(* IEC 61131-3 sources: plc-vscode/tests/st/test-ready/rusty/tests/lit/single/polymorphism/properties, 4 files *)

(* ---- alternating_accessor_overrides.st ---- *)
// RUN: (%COMPILE %s && %RUN) | %CHECK %s
// Scenario: Three-level POU chain C → B → A. B overrides only the getter (adds 1000),
// C overrides only the setter (adds 2000). Dispatch through POINTER TO A should resolve
// each accessor independently to the most-derived override:
//   A → (A.get, A.set)
//   B → (B.get, A.set)
//   C → (B.get, C.set)

FUNCTION_BLOCK A
    VAR
        _val : DINT := 10;
    END_VAR

    PROPERTY_GET value: DINT
        value := _val;
    END_PROPERTY

    PROPERTY_SET value: DINT
        _val := value;
    END_PROPERTY

    METHOD printValue
        printf('value=%d$N', value);
    END_METHOD

    METHOD setValue
        VAR_INPUT x : DINT; END_VAR
        value := x;
    END_METHOD
END_FUNCTION_BLOCK

FUNCTION_BLOCK B EXTENDS A
    // Override only getter — adds 1000
    PROPERTY_GET value: DINT
        value := _val + 1000;
    END_PROPERTY
END_FUNCTION_BLOCK

FUNCTION_BLOCK C EXTENDS B
    // Override only setter — adds 2000
    PROPERTY_SET value: DINT
        _val := value + 2000;
    END_PROPERTY
END_FUNCTION_BLOCK

FUNCTION printViaPtr
    VAR_INPUT
        p : POINTER TO A;
    END_VAR

    p^.printValue();
END_FUNCTION

FUNCTION setViaPtr
    VAR_INPUT
        p : POINTER TO A;
        x : DINT;
    END_VAR

    p^.setValue(x);
END_FUNCTION

FUNCTION main
    VAR
        instanceA : A;
        instanceB : B;
        instanceC : C;
    END_VAR

    // A: get=A, set=A
    printViaPtr(ADR(instanceA));        // CHECK: value=10
    setViaPtr(ADR(instanceA), 50);
    printViaPtr(ADR(instanceA));        // CHECK-NEXT: value=50

    // B: get=B(+1000), set=A(inherited)
    printViaPtr(ADR(instanceB));        // CHECK-NEXT: value=1010
    setViaPtr(ADR(instanceB), 50);
    printViaPtr(ADR(instanceB));        // CHECK-NEXT: value=1050

    // C: get=B(inherited, +1000), set=C(+2000)
    printViaPtr(ADR(instanceC));        // CHECK-NEXT: value=1010
    setViaPtr(ADR(instanceC), 50);
    printViaPtr(ADR(instanceC));        // CHECK-NEXT: value=3050
END_FUNCTION

(* ---- inherited_getter_overridden_setter.st ---- *)
// RUN: (%COMPILE %s && %RUN) | %CHECK %s
// Scenario: B extends A which has a property with both PROPERTY_GET and PROPERTY_SET. B overrides only the setter.
// Dispatch through POINTER TO A should use A's inherited getter and B's overridden setter.

FUNCTION_BLOCK A
    VAR
        _val : DINT := 10;
    END_VAR

    PROPERTY_GET value: DINT
        value := _val;
    END_PROPERTY

    PROPERTY_SET value: DINT
        _val := value;
    END_PROPERTY

    METHOD printValue
        printf('value=%d$N', value);
    END_METHOD

    METHOD setValue
        VAR_INPUT x : DINT; END_VAR
        value := x;
    END_METHOD
END_FUNCTION_BLOCK

FUNCTION_BLOCK B EXTENDS A
    // Override only the setter — adds 1000 to distinguish from A's setter
    PROPERTY_SET value: DINT
        _val := value + 1000;
    END_PROPERTY
END_FUNCTION_BLOCK

FUNCTION printViaPtr
    VAR_INPUT
        p : POINTER TO A;
    END_VAR

    p^.printValue();
END_FUNCTION

FUNCTION setViaPtr
    VAR_INPUT
        p : POINTER TO A;
        x : DINT;
    END_VAR

    p^.setValue(x);
END_FUNCTION

FUNCTION main
    VAR
        instanceA : A;
        instanceB : B;
    END_VAR

    // A — base getter and setter
    printViaPtr(ADR(instanceA));        // CHECK: value=10
    setViaPtr(ADR(instanceA), 42);
    printViaPtr(ADR(instanceA));        // CHECK-NEXT: value=42

    // B — inherited getter, overridden setter (adds 1000)
    printViaPtr(ADR(instanceB));        // CHECK-NEXT: value=10
    setViaPtr(ADR(instanceB), 42);
    printViaPtr(ADR(instanceB));        // CHECK-NEXT: value=1042
END_FUNCTION

(* ---- method_dispatches_to_overridden_property.st ---- *)
// RUN: (%COMPILE %s && %RUN) | %CHECK %s
// Scenario: A defines a method `doubleValue` that reads and writes a property internally.
// B extends A and overrides only the setter (adds 100). When `doubleValue` is called on a B
// instance through POINTER TO A, the read dispatches to A's getter but the write dispatches
// to B's overridden setter — proving that property dispatch inside a non-overridden method
// is truly dynamic.

FUNCTION_BLOCK A
    VAR
        _val : DINT := 5;
    END_VAR

    PROPERTY_GET value: DINT
        value := _val;
    END_PROPERTY

    PROPERTY_SET value: DINT
        _val := value;
    END_PROPERTY

    METHOD doubleValue
        value := value * 2;
    END_METHOD

    METHOD printValue
        printf('value=%d$N', value);
    END_METHOD
END_FUNCTION_BLOCK

FUNCTION_BLOCK B EXTENDS A
    // Override only setter — adds 100
    PROPERTY_SET value: DINT
        _val := value + 100;
    END_PROPERTY
END_FUNCTION_BLOCK

FUNCTION printViaPtr
    VAR_INPUT
        p : POINTER TO A;
    END_VAR

    p^.printValue();
END_FUNCTION

FUNCTION doubleViaPtr
    VAR_INPUT
        p : POINTER TO A;
    END_VAR

    p^.doubleValue();
END_FUNCTION

FUNCTION main
    VAR
        instanceA : A;
        instanceB : B;
    END_VAR

    // A — base: doubleValue reads 5, writes 10
    printViaPtr(ADR(instanceA));        // CHECK: value=5
    doubleViaPtr(ADR(instanceA));
    printViaPtr(ADR(instanceA));        // CHECK-NEXT: value=10
    doubleViaPtr(ADR(instanceA));
    printViaPtr(ADR(instanceA));        // CHECK-NEXT: value=20

    // B — inherited getter, overridden setter (+100)
    // doubleValue reads 5 (A.get), writes 10 → B.set stores 10+100=110
    printViaPtr(ADR(instanceB));        // CHECK-NEXT: value=5
    doubleViaPtr(ADR(instanceB));
    printViaPtr(ADR(instanceB));        // CHECK-NEXT: value=110
    // doubleValue reads 110 (A.get), writes 220 → B.set stores 220+100=320
    doubleViaPtr(ADR(instanceB));
    printViaPtr(ADR(instanceB));        // CHECK-NEXT: value=320
END_FUNCTION

(* ---- multiple_properties_selective_overrides.st ---- *)
// RUN: (%COMPILE %s && %RUN) | %CHECK %s
// Scenario: A has two properties (x and y). B extends A and overrides only the getter of x
// (adds 100) and only the setter of y (adds 200). Dispatch through POINTER TO A verifies
// that each property's each accessor is resolved independently through the vtable.

FUNCTION_BLOCK A
    VAR
        _x : DINT := 1;
        _y : DINT := 2;
    END_VAR

    PROPERTY_GET x: DINT
        x := _x;
    END_PROPERTY

    PROPERTY_SET x: DINT
        _x := x;
    END_PROPERTY

    PROPERTY_GET y: DINT
        y := _y;
    END_PROPERTY

    PROPERTY_SET y: DINT
        _y := y;
    END_PROPERTY

    METHOD printXY
        printf('x=%d, y=%d$N', x, y);
    END_METHOD

    METHOD setX
        VAR_INPUT v : DINT; END_VAR
        x := v;
    END_METHOD

    METHOD setY
        VAR_INPUT v : DINT; END_VAR
        y := v;
    END_METHOD
END_FUNCTION_BLOCK

FUNCTION_BLOCK B EXTENDS A
    // Override only getter of x — adds 100
    PROPERTY_GET x: DINT
        x := _x + 100;
    END_PROPERTY

    // Override only setter of y — adds 200
    PROPERTY_SET y: DINT
        _y := y + 200;
    END_PROPERTY
END_FUNCTION_BLOCK

FUNCTION printViaPtr
    VAR_INPUT
        p : POINTER TO A;
    END_VAR

    p^.printXY();
END_FUNCTION

FUNCTION setXViaPtr
    VAR_INPUT
        p : POINTER TO A;
        v : DINT;
    END_VAR

    p^.setX(v);
END_FUNCTION

FUNCTION setYViaPtr
    VAR_INPUT
        p : POINTER TO A;
        v : DINT;
    END_VAR

    p^.setY(v);
END_FUNCTION

FUNCTION main
    VAR
        instanceA : A;
        instanceB : B;
    END_VAR

    // A: x.get=A, x.set=A, y.get=A, y.set=A
    printViaPtr(ADR(instanceA));                // CHECK: x=1, y=2
    setXViaPtr(ADR(instanceA), 10);
    setYViaPtr(ADR(instanceA), 20);
    printViaPtr(ADR(instanceA));                // CHECK-NEXT: x=10, y=20

    // B: x.get=B(+100), x.set=A(inherited), y.get=A(inherited), y.set=B(+200)
    printViaPtr(ADR(instanceB));                // CHECK-NEXT: x=101, y=2
    setXViaPtr(ADR(instanceB), 10);
    setYViaPtr(ADR(instanceB), 20);
    printViaPtr(ADR(instanceB));                // CHECK-NEXT: x=110, y=220
END_FUNCTION
